# EPICS StreamDevice protocol: reference/lab-2023/EPICS/Db/aim.proto
# Author: Philip Weigel

Terminator = CR;

get_pressure {
	out "?V752";
	in "=V752 %E;%*d";
}

enable {
	out "\!C752 %{0|1}";
}
